(* IEC 61131-3 sources: iolistgen/tests_support/pl_stub/src/DUTs/Alarm, 5 files *)

(* ---- E_AlarmEventReason.dut.st ---- *)
// Назначение: заглушка plc-process-lib 1.0.0 для проверки типов сгенерированного кода без CODESYS
//             (API.md, раздел 4.1); не библиотека — тел и внутренних переменных нет
// Автор:      kr0nsch
// Версия:     1.0.0 (выпуск библиотеки)
// Документ:   docs/GENERATORS.md, раздел «Проверка ST без CODESYS»
{attribute 'qualified_only'}
{attribute 'strict'}
TYPE E_AlarmEventReason :
(
    None := 0,
    Activated := 1,
    Cleared := 2,
    Acked := 3,
    Shelved := 4,
    Unshelved := 5,
    ShelveExpired := 6,
    Suppressed := 7,
    Unsuppressed := 8,
    OosOn := 9,
    OosOff := 10,
    Disabled := 11
) INT;
END_TYPE

(* ---- E_AlarmPriority.dut.st ---- *)
// Назначение: заглушка plc-process-lib 1.0.0 для проверки типов сгенерированного кода без CODESYS
//             (API.md, раздел 4.1); не библиотека — тел и внутренних переменных нет
// Автор:      kr0nsch
// Версия:     1.0.0 (выпуск библиотеки)
// Документ:   docs/GENERATORS.md, раздел «Проверка ST без CODESYS»
{attribute 'qualified_only'}
{attribute 'strict'}
TYPE E_AlarmPriority :
(
    None := 0,
    Low := 1,
    Medium := 2,
    High := 3,
    Critical := 4
) INT;
END_TYPE

(* ---- E_AlarmState.dut.st ---- *)
// Назначение: заглушка plc-process-lib 1.0.0 для проверки типов сгенерированного кода без CODESYS
//             (API.md, раздел 4.1); не библиотека — тел и внутренних переменных нет
// Автор:      kr0nsch
// Версия:     1.0.0 (выпуск библиотеки)
// Документ:   docs/GENERATORS.md, раздел «Проверка ST без CODESYS»
{attribute 'qualified_only'}
{attribute 'strict'}
TYPE E_AlarmState :
(
    Normal := 0,
    ActiveUnack := 1,
    ActiveAck := 2,
    RtnUnack := 3,
    Shelved := 4,
    SuppressedByDesign := 5,
    OutOfService := 6
) INT;
END_TYPE

(* ---- ST_AlarmCfg.dut.st ---- *)
// Назначение: заглушка plc-process-lib 1.0.0 для проверки типов сгенерированного кода без CODESYS
//             (API.md, раздел 4.4); не библиотека — тел и внутренних переменных нет
// Автор:      kr0nsch
// Версия:     1.0.0 (выпуск библиотеки)
// Документ:   docs/GENERATORS.md, раздел «Проверка ST без CODESYS»
{attribute 'qualified_only'}
TYPE ST_AlarmCfg :
STRUCT
    ePriority  : E_AlarmPriority := E_AlarmPriority.Medium;
    tOnDelay   : TIME := T#0S;
    tOffDelay  : TIME := T#0S;
    tShelveMax : TIME := T#8H;
END_STRUCT
END_TYPE

(* ---- ST_AlarmEvent.dut.st ---- *)
// Назначение: заглушка plc-process-lib 1.0.0 для проверки типов сгенерированного кода без CODESYS
//             (API.md, раздел 4.4); не библиотека — тел и внутренних переменных нет
// Автор:      kr0nsch
// Версия:     1.0.0 (выпуск библиотеки)
// Документ:   docs/GENERATORS.md, раздел «Проверка ST без CODESYS»
{attribute 'qualified_only'}
TYPE ST_AlarmEvent :
STRUCT
    udiId     : UDINT;
    ePriority : E_AlarmPriority;
    eOldState : E_AlarmState;
    eNewState : E_AlarmState;
    eReason   : E_AlarmEventReason;
    ltTime    : LTIME;
    rValue    : REAL;
END_STRUCT
END_TYPE
